Staubli VAL3: stop.pgx

program stop()
begin
  //应用停止时调用：让机器人停在安全状态
  bRunning=false
  nState=0
end
